TYPE ST_ReadBlock :
STRUCT
    startAddress        : UINT;
    quantity            : UINT;
    area                : E_MBArea;
    functionCode        : BYTE;

    arrSignalIndex      : ARRAY[1..64] OF UINT;
    arrOffsetInBlock    : ARRAY[1..64] OF UINT;
    signalCount         : UINT;

    enabled             : BOOL := TRUE;
END_STRUCT
END_TYPE

(* stored: Version 1.1.0.1, ProductVersion 3.1.4024.0
   DUT ST_ReadBlock: Id {3401096d-414a-42f9-9e85-c401026e9f45} *)
